(* IEC 61131-3 sources: llm-plc-st-eval/data/processed_definitivo/claude-sonnet-4-6/A6/few_shot, 3 files *)

(* ---- ejec_1.st ---- *)
FUNCTION_BLOCK FB_Modos
VAR_INPUT
    selector       : INT;                  (* Selector de modo: 0=Auto, 1=Manual, 2=Mantenimiento *)
    estadoSeguro   : BOOL;                 (* Permiso para cambiar de modo y operar mantenimiento *)
    cmdAuto        : ARRAY[0..7] OF BOOL;  (* Comandos en modo automatico *)
    cmdManual      : ARRAY[0..7] OF BOOL;  (* Comandos en modo manual *)
    idxForzado     : INT;                  (* Indice del actuador a forzar en mantenimiento *)
    valorForzado   : BOOL;                 (* Valor a aplicar al actuador forzado *)
    confirmarForzado : BOOL;               (* Flanco ascendente aplica el forzado *)
END_VAR
VAR_OUTPUT
    modoActivo : INT;                      (* Modo vigente: 0=Auto, 1=Manual, 2=Mantenimiento *)
    actuador   : ARRAY[0..7] OF BOOL;      (* Estado de los ocho actuadores *)
END_VAR
VAR
    prevConfirmar  : BOOL;                 (* Valor anterior de confirmarForzado para deteccion de flanco *)
    estadoForzado  : ARRAY[0..7] OF BOOL;  (* Valores forzados en modo mantenimiento *)
    i              : INT;                  (* Indice auxiliar para bucles *)
    primerCiclo    : BOOL := TRUE;         (* Marca de primer ciclo para inicializacion *)
END_VAR

(* --- Inicializacion en el primer ciclo de ejecucion --- *)
IF primerCiclo THEN
    modoActivo  := 1;   (* Modo inicial: manual *)
    primerCiclo := FALSE;
END_IF;

(* --- Gestion del cambio de modo --- *)
(* Solo se acepta un nuevo modo si estadoSeguro esta activo y el valor es valido (0..2) *)
IF estadoSeguro AND (selector >= 0) AND (selector <= 2) THEN
    IF selector <> modoActivo THEN
        (* Al salir del modo mantenimiento se anulan todos los forzados *)
        IF modoActivo = 2 THEN
            FOR i := 0 TO 7 DO
                estadoForzado[i] := FALSE;
            END_FOR;
        END_IF;
        modoActivo := selector;
    END_IF;
END_IF;

(* --- Logica especifica de cada modo --- *)
CASE modoActivo OF

    0: (* Modo automatico: actuadores siguen cmdAuto *)
        FOR i := 0 TO 7 DO
            actuador[i] := cmdAuto[i];
        END_FOR;

    1: (* Modo manual: actuadores siguen cmdManual *)
        FOR i := 0 TO 7 DO
            actuador[i] := cmdManual[i];
        END_FOR;

    2: (* Modo mantenimiento *)
        IF NOT estadoSeguro THEN
            (* Si se pierde el estado seguro, se anulan forzados y se apagan actuadores *)
            FOR i := 0 TO 7 DO
                estadoForzado[i] := FALSE;
                actuador[i]      := FALSE;
            END_FOR;
        ELSE
            (* Deteccion de flanco ascendente en confirmarForzado *)
            IF confirmarForzado AND NOT prevConfirmar THEN
                IF (idxForzado >= 0) AND (idxForzado <= 7) THEN
                    estadoForzado[idxForzado] := valorForzado;
                END_IF;
                (* Indices fuera de rango se ignoran *)
            END_IF;
            (* Los actuadores reflejan el estado forzado acumulado *)
            FOR i := 0 TO 7 DO
                actuador[i] := estadoForzado[i];
            END_FOR;
        END_IF;

END_CASE;

(* --- Actualizacion del valor previo de confirmarForzado --- *)
prevConfirmar := confirmarForzado;

END_FUNCTION_BLOCK

(* ---- ejec_2.st ---- *)
FUNCTION_BLOCK FB_Modos
VAR_INPUT
    selector       : INT;                  (* Selector de modo: 0=Auto, 1=Manual, 2=Mantenimiento *)
    estadoSeguro   : BOOL;                 (* Permiso para cambiar modo y mantener forzados *)
    cmdAuto        : ARRAY[0..7] OF BOOL;  (* Comandos en modo automatico *)
    cmdManual      : ARRAY[0..7] OF BOOL;  (* Comandos en modo manual *)
    idxForzado     : INT;                  (* Indice del actuador a forzar (0..7) *)
    valorForzado   : BOOL;                 (* Valor a aplicar al actuador forzado *)
    confirmarForzado : BOOL;               (* Flanco ascendente aplica el forzado *)
END_VAR
VAR_OUTPUT
    modoActivo : INT;                      (* Modo vigente: 0=Auto, 1=Manual, 2=Mantenimiento *)
    actuador   : ARRAY[0..7] OF BOOL;      (* Estado de los ocho actuadores *)
END_VAR
VAR
    modoInterno        : INT := 1;         (* Modo interno; arranca en manual *)
    estadoSeguroPrev   : BOOL;             (* Valor anterior de estadoSeguro *)
    confirmarForzadoPrev : BOOL;           (* Valor anterior de confirmarForzado para deteccion de flanco *)
    estadoForzado      : ARRAY[0..7] OF BOOL; (* Valores forzados en mantenimiento *)
    i                  : INT;             (* Indice de iteracion *)
    primeraEjecucion   : BOOL := TRUE;    (* Bandera de primera ejecucion *)
END_VAR

(* --- Inicializacion en primera ejecucion --- *)
IF primeraEjecucion THEN
    modoInterno      := 1; (* Manual por defecto *)
    primeraEjecucion := FALSE;
END_IF;

(* --- Gestion de cambio de modo --- *)
(* Solo se acepta un nuevo modo si estadoSeguro esta activo y el valor es valido (0..2) *)
IF estadoSeguro AND (selector >= 0) AND (selector <= 2) AND (selector <> modoInterno) THEN
    (* Al salir de mantenimiento, anular todos los forzados *)
    IF modoInterno = 2 THEN
        FOR i := 0 TO 7 DO
            estadoForzado[i] := FALSE;
        END_FOR;
    END_IF;
    modoInterno := selector;
END_IF;

(* --- Deteccion de flanco descendente en estadoSeguro durante mantenimiento --- *)
(* Si estadoSeguro se desactiva en modo mantenimiento, apagar todos los actuadores forzados *)
IF (NOT estadoSeguro) AND estadoSeguroPrev AND (modoInterno = 2) THEN
    FOR i := 0 TO 7 DO
        estadoForzado[i] := FALSE;
    END_FOR;
END_IF;
estadoSeguroPrev := estadoSeguro;

(* --- Logica segun modo activo --- *)
CASE modoInterno OF

    0: (* Modo automatico: actuadores siguen cmdAuto *)
        FOR i := 0 TO 7 DO
            actuador[i] := cmdAuto[i];
        END_FOR;

    1: (* Modo manual: actuadores siguen cmdManual *)
        FOR i := 0 TO 7 DO
            actuador[i] := cmdManual[i];
        END_FOR;

    2: (* Modo mantenimiento *)
        (* Forzado individual con flanco ascendente de confirmarForzado *)
        (* Solo se procesa si estadoSeguro esta activo *)
        IF estadoSeguro AND confirmarForzado AND (NOT confirmarForzadoPrev) THEN
            IF (idxForzado >= 0) AND (idxForzado <= 7) THEN
                estadoForzado[idxForzado] := valorForzado;
            END_IF;
        END_IF;
        (* Los actuadores reflejan el estado forzado *)
        FOR i := 0 TO 7 DO
            actuador[i] := estadoForzado[i];
        END_FOR;

END_CASE;

(* --- Actualizar flanco de confirmarForzado --- *)
confirmarForzadoPrev := confirmarForzado;

(* --- Reportar modo vigente --- *)
modoActivo := modoInterno;

END_FUNCTION_BLOCK

(* ---- ejec_3.st ---- *)
FUNCTION_BLOCK FB_Modos
VAR_INPUT
    selector       : INT;                  (* Selector de modo: 0=Auto, 1=Manual, 2=Mant. *)
    estadoSeguro   : BOOL;                 (* Permiso para cambio de modo y forzados *)
    cmdAuto        : ARRAY[0..7] OF BOOL;  (* Comandos en modo automatico *)
    cmdManual      : ARRAY[0..7] OF BOOL;  (* Comandos en modo manual *)
    idxForzado     : INT;                  (* Indice del actuador a forzar (0..7) *)
    valorForzado   : BOOL;                 (* Valor a aplicar al actuador forzado *)
    confirmarForzado : BOOL;               (* Flanco ascendente aplica el forzado *)
END_VAR
VAR_OUTPUT
    modoActivo : INT;                      (* Modo vigente: 0=Auto, 1=Manual, 2=Mant. *)
    actuador   : ARRAY[0..7] OF BOOL;     (* Estado de los ocho actuadores *)
END_VAR
VAR
    i                  : INT;             (* Indice de bucle *)
    estadosForzados    : ARRAY[0..7] OF BOOL; (* Valores forzados en mantenimiento *)
    confirmarForzado_prev : BOOL;         (* Valor anterior de confirmarForzado *)
    flanco_confirmar   : BOOL;            (* Flanco ascendente detectado *)
    primerCiclo        : BOOL := TRUE;    (* Bandera de primer ciclo para inicializacion *)
    estadoSeguro_prev  : BOOL;            (* Valor anterior de estadoSeguro *)
END_VAR

(* --- Inicializacion en el primer ciclo: modo manual por defecto --- *)
IF primerCiclo THEN
    modoActivo        := 1;
    primerCiclo       := FALSE;
    confirmarForzado_prev := confirmarForzado;
    estadoSeguro_prev := estadoSeguro;
    FOR i := 0 TO 7 DO
        estadosForzados[i] := FALSE;
        actuador[i]        := FALSE;
    END_FOR;
END_IF;

(* --- Gestion del cambio de modo --- *)
(* Solo se acepta un selector valido (0..2) y con estadoSeguro activo *)
IF estadoSeguro AND (selector >= 0) AND (selector <= 2) THEN
    IF selector <> modoActivo THEN
        (* Al salir de mantenimiento, anular todos los forzados *)
        IF modoActivo = 2 THEN
            FOR i := 0 TO 7 DO
                estadosForzados[i] := FALSE;
            END_FOR;
        END_IF;
        modoActivo := selector;
        (* Al entrar en mantenimiento, apagar todos los actuadores *)
        IF modoActivo = 2 THEN
            FOR i := 0 TO 7 DO
                actuador[i]        := FALSE;
                estadosForzados[i] := FALSE;
            END_FOR;
        END_IF;
    END_IF;
END_IF;

(* --- Logica especifica de mantenimiento --- *)
IF modoActivo = 2 THEN
    (* Si estadoSeguro se desactiva durante mantenimiento: anular forzados y apagar *)
    IF (NOT estadoSeguro) AND estadoSeguro_prev THEN
        FOR i := 0 TO 7 DO
            estadosForzados[i] := FALSE;
            actuador[i]        := FALSE;
        END_FOR;
    END_IF;

    (* Detectar flanco ascendente de confirmarForzado *)
    flanco_confirmar := confirmarForzado AND (NOT confirmarForzado_prev);

    (* Aplicar forzado solo si estadoSeguro activo, flanco detectado e indice valido *)
    IF estadoSeguro AND flanco_confirmar
       AND (idxForzado >= 0) AND (idxForzado <= 7) THEN
        estadosForzados[idxForzado] := valorForzado;
    END_IF;

    (* Los actuadores reflejan los valores forzados *)
    FOR i := 0 TO 7 DO
        actuador[i] := estadosForzados[i];
    END_FOR;

(* --- Modo automatico --- *)
ELSIF modoActivo = 0 THEN
    FOR i := 0 TO 7 DO
        actuador[i] := cmdAuto[i];
    END_FOR;

(* --- Modo manual --- *)
ELSIF modoActivo = 1 THEN
    FOR i := 0 TO 7 DO
        actuador[i] := cmdManual[i];
    END_FOR;
END_IF;

(* --- Actualizar valores previos para el proximo ciclo --- *)
confirmarForzado_prev := confirmarForzado;
estadoSeguro_prev     := estadoSeguro;

END_FUNCTION_BLOCK
